(* IEC 61131-3 sources: codesys-to-astra/corpus/boiler-plc210/src/POUs/PRG_Slow, 2 files *)

(* ---- PRG_Slow.decl.st ---- *)
// Назначение: медленная задача (приоритет 15 у ОВЕН): слово состояния панели.
// Автор:      kr0nsch
// Версия:     0.1.0
// Документ:   corpus/boiler-plc210/README.md
PROGRAM PRG_Slow
VAR
END_VAR
VAR CONSTANT
    BIT_FAULT : WORD := 16#0002;    // бит «авария» в слове состояния
    BIT_RUN : WORD := 16#0001;      // бит «работа»
END_VAR

(* ---- PRG_Slow.impl.st ---- *)
GVL_Hw.wHmiStatus := 0;
IF GVL_Hmi.eState = E_BoilerState.Run THEN
    GVL_Hw.wHmiStatus := GVL_Hw.wHmiStatus OR BIT_RUN;
END_IF
IF GVL_Hmi.eState = E_BoilerState.Fault THEN
    GVL_Hw.wHmiStatus := GVL_Hw.wHmiStatus OR BIT_FAULT;
END_IF
